Staubli VAL3: insertFOR.pgx

public program insertFOR(num x_nProgIndex)
  local bool l_bExit
  local bool l_bRefreh
  local num l_nProgIndex
  local num l_i
  local bool l_bRefresh
begin
  do
    if util:sPage!="insertFOR"
      util:sPage="insertFOR"
      call _onStartPROG(util:sPage)
      call _bindPROG(util:sPage)
      userPageBind("insertFOR","nmb1","value",nFORValue,1,"rw")
      if size(sIOList)!=(size(io:aInItem)+1)
        resize(sIOList,1,size(io:aInItem)+1)
      endIf
      for l_i = 1 to size(sIOList)-1
        sIOList[l_i-1]=toString("",l_i-1)+","+io:aInItem[l_i-1].sComment
      endFor
      sIOList[0]="value"
      userPageBind("insertFOR","cbx1","options",sIOList,size(sIOList),"r")
      userPageBind("insertFOR","cbx1","value",sForValue,1,"rw")
      userPage(util:sPage)
      delay(0.5)
    endIf

    //btn
    if bSelProg
      bSelProg=false
      nSelType=1
      l_bRefresh=true
      nPgIndexPROG=0
    elseIf bSelTraj
      bSelTraj=false
      nSelType=2
      l_bRefresh=true
      nPgIndexPROG=0
    endIf


    //refresh
    if l_bRefresh
      l_bRefresh=false
      call _btnColor(nSelType,util:sPage)
      switch nSelType
        case 1
          call resfreshPROG(util:sPage)
        break
        case 2
          nPgIndexTRAJ=0
          call resfreshTRAJ(util:sPage)
        break
      endSwitch
    endIf

    if bInsert[1]
      bInsert[1]=false

      call prog:insertFOR(sSelProg,x_nProgIndex,sInsertItem,nFORValue,sForValue,bToSave,nSelType)

      l_bExit=true
    elseIf bInsert[2]
      bInsert[2]=false
      l_bExit=true
    elseIf bInsert[3]
      bInsert[3]=false
      nPgIndexPROG=0
      l_bRefreh=true
    elseIf bInsert[4]
      bInsert[4]=false
      if nPgIndexPROG>0
        nPgIndexPROG=nPgIndexPROG-1
        l_bRefreh=true
      endIf

    elseIf bInsert[5]
      bInsert[5]=false
      if nPgIndexPROG<nPgNumPROG-1
        nPgIndexPROG=nPgIndexPROG+1
        l_bRefreh=true
      endIf

    elseIf bInsert[6]
      bInsert[6]=false
      nPgIndexPROG=nPgNumPROG-1
      l_bRefreh=true
    endIf





    delay(0)
  until l_bExit==true
end
